FUNCTION_BLOCK FB_ReversibleConveyor EXTENDS FB_ConveyorBase IMPLEMENTS I_Reversible
VAR
    reverseState : BOOL;
END_VAR

PROPERTY PUBLIC Reverse : BOOL
GET
Reverse := reverseState;
END_GET
SET
reverseState := Reverse;
END_SET
END_PROPERTY

PROPERTY PUBLIC ActualSpeed : REAL
GET
ActualSpeed := SUPER^.ActualSpeed;
IF reverseState THEN ActualSpeed := -ActualSpeed; END_IF;
END_GET
END_PROPERTY

END_FUNCTION_BLOCK

(* stored: Version 1.1.0.1, ProductVersion 3.1 *)
